Fanuc KAREL source: KD00012.KL

PROGRAM KD00012
%NOLOCKGROUP
VAR
  I: INTEGER
  J: INTEGER
  B: BOOLEAN
  R: REAL
  S: STRING[80]
BEGIN
  OPEN HAND 1
END KD00012
